// TIA Portal V19 export
FUNCTION_BLOCK "MOTOR"   // FB4, FBD
{ S7_Optimized_Access := 'TRUE' }
// stored: MemoryReserve 100, SetENOAutomatically false
   VAR
      AG_01 { S7_SetPoint := 'True'} : "MOTOR_FB1";
   END_VAR
BEGIN

REGION Network 1: Agitator
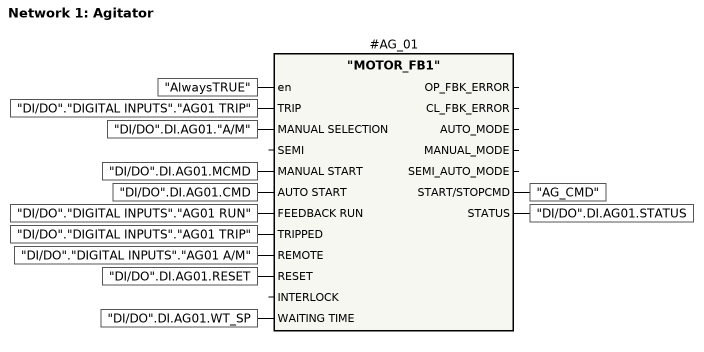
   IF "AlwaysTRUE" THEN
       #AG_01(TRIP := "DI/DO"."DIGITAL INPUTS"."AG01 TRIP",   // "MOTOR_FB1"
              "MANUAL SELECTION" := "DI/DO".DI.AG01."A/M",
              "MANUAL START" := "DI/DO".DI.AG01.MCMD,
              "AUTO START" := "DI/DO".DI.AG01.CMD,
              "FEEDBACK RUN" := "DI/DO"."DIGITAL INPUTS"."AG01 RUN",
              TRIPPED := "DI/DO"."DIGITAL INPUTS"."AG01 TRIP",
              REMOTE := "DI/DO"."DIGITAL INPUTS"."AG01 A/M",
              RESET := "DI/DO".DI.AG01.RESET,
              "WAITING TIME" := "DI/DO".DI.AG01.WT_SP,
              "START/STOPCMD" => "AG_CMD",
              STATUS => "DI/DO".DI.AG01.STATUS);
   END_IF;
END_REGION
END_FUNCTION_BLOCK
